(* CODESYS project getsystemtime.library
   DefaultNamespace: KOSTAL.AF2024.Core.GetSystemTime
   DocFormat: reStructuredText
   Description: Contains Functionalities to get the NT Real Time Clock
   Author: Frank Dümpelmann
   Title: KOSTAL.AF2024.Core.GetSystemTime
   Version: 1.0.1.0
   Company: KOSTAL GmbH & Co.KG
   Placeholder: KOSTAL.AF2024.Core.GetSystemTime

Project tree, tasks and I/O mapping:
  libraries: Tc2_Utilities, 3.3.47.0 (Beckhoff Automation GmbH); KOSTAL.AF2024.Core.System, 1.0.0.0 (KOSTAL GmbH & Co.KG)
  DUT/
    data type E_TIMESHIFT
    interface I_T_Timestruct: CopyTo, Day, DayOfWeek, Hour, iTimeStruct, Milliseconds, Minute, Month, Second, Year
    interface I_T_Timestruct_Owner: Day, DayOfWeek, Hour, Milliseconds, Minute, Month, Second, Timestruct, Year
    data type ST_TIMEZONE
    function block T_TIMESTRUCT [ST]: CopyTo, Day, DayOfWeek, Hour, iTimeStruct, Milliseconds, Minute, Month, Second, Timestruct, Year
  Interface/
    interface I_TimeSource: DateAndTime, GetTimeStruct, GetTimeZone, TimeStruct, Utc, Valid
  POU/
    function block FB_GetSystemTime [ST]: _formatTimeZone, amsNetId_timeServer, DateAndTime, FBmain, GetTimeStruct, GetTimeZone, Timeout, TimeStruct, Utc, Valid
  Project Information/
    function F_GetCompany [ST]
    function F_GetTitle [ST]
    function F_GetVersion [ST]
  Version/
    global variables Global_Version
*)

// DUT/E_TIMESHIFT
{attribute 'qualified_only'}
{attribute 'strict'}
TYPE E_TIMESHIFT :
(
	undef 		:= 0,
	positive 	:= 1,
	negative 	:= 2
);
END_TYPE

// DUT/ST_TIMEZONE
TYPE ST_TIMEZONE :
STRUCT
	timeshift	: E_TIMESHIFT;
	hours		: USINT;
	minutes		: USINT;
END_STRUCT
END_TYPE

// Version/Global_Version
{attribute 'TcGenerated'}
{attribute 'no-analysis'}
{attribute 'linkalways'}
// This function has been automatically generated from the project information.
VAR_GLOBAL CONSTANT
	{attribute 'const_non_replaced'}
	stLibVersion_KOSTAL_AF2024_Core_GetSystemTime : ST_LibVersion := (iMajor := 1, iMinor := 0, iBuild := 1, iRevision := 0, nFlags := 1, sVersion := '1.0.1.0');
END_VAR

// DUT/I_T_Timestruct
INTERFACE I_T_Timestruct EXTENDS KOSTAL_AF2024_Core_System.I_Interface

METHOD CopyTo
VAR_INPUT
	IN : REFERENCE TO Tc2_Utilities.TIMESTRUCT;
END_VAR
END_METHOD

PROPERTY PUBLIC Day : WORD
GET
END_GET
END_PROPERTY

PROPERTY PUBLIC DayOfWeek : WORD
GET
END_GET
END_PROPERTY

PROPERTY PUBLIC Hour : WORD
GET
END_GET
END_PROPERTY

PROPERTY iTimeStruct : Tc2_Utilities.TIMESTRUCT
GET
END_GET
END_PROPERTY

PROPERTY PUBLIC Milliseconds : WORD
GET
END_GET
END_PROPERTY

PROPERTY PUBLIC Minute : WORD
GET
END_GET
END_PROPERTY

PROPERTY PUBLIC Month : WORD
GET
END_GET
END_PROPERTY

PROPERTY PUBLIC Second : WORD
GET
END_GET
END_PROPERTY

PROPERTY PUBLIC Year : WORD
GET
END_GET
END_PROPERTY

END_INTERFACE

// DUT/I_T_Timestruct_Owner
INTERFACE I_T_Timestruct_Owner EXTENDS KOSTAL_AF2024_Core_System.I_Interface

PROPERTY PUBLIC Day : WORD
GET
END_GET
SET
END_SET
END_PROPERTY

PROPERTY PUBLIC DayOfWeek : WORD
GET
END_GET
SET
END_SET
END_PROPERTY

PROPERTY PUBLIC Hour : WORD
GET
END_GET
SET
END_SET
END_PROPERTY

PROPERTY PUBLIC Milliseconds : WORD
GET
END_GET
SET
END_SET
END_PROPERTY

PROPERTY PUBLIC Minute : WORD
GET
END_GET
SET
END_SET
END_PROPERTY

PROPERTY PUBLIC Month : WORD
GET
END_GET
SET
END_SET
END_PROPERTY

PROPERTY PUBLIC Second : WORD
GET
END_GET
SET
END_SET
END_PROPERTY

PROPERTY Timestruct : REFERENCE To Tc2_Utilities.TIMESTRUCT
GET
END_GET
END_PROPERTY

PROPERTY PUBLIC Year : WORD
GET
END_GET
SET
END_SET
END_PROPERTY

END_INTERFACE

// DUT/T_TIMESTRUCT
FUNCTION_BLOCK T_TIMESTRUCT IMPLEMENTS I_T_Timestruct, I_T_Timestruct_Owner
VAR
	_timestruct : Tc2_Utilities.TIMESTRUCT;
END_VAR

METHOD CopyTo
VAR_INPUT
	IN : REFERENCE TO Tc2_Utilities.TIMESTRUCT;
END_VAR

IN.wYear := _timestruct.wYear;
IN.wMonth := _timestruct.wMonth;
IN.wDay := _timestruct.wDay;
IN.wDayOfWeek := _timestruct.wDayOfWeek;
IN.wHour := _timestruct.wHour;
IN.wMinute := _timestruct.wMinute;
IN.wSecond := _timestruct.wSecond;
IN.wMilliseconds := _timestruct.wMilliseconds;
END_METHOD

PROPERTY PUBLIC Day : WORD
GET
Day := _timestruct.wDay;
END_GET
SET
_timestruct.wDay := Day;
END_SET
END_PROPERTY

PROPERTY PUBLIC DayOfWeek : WORD
GET
DayOfWeek := _timestruct.wDayOfWeek;
END_GET
SET
_timestruct.wDayOfWeek := DayOfWeek;
END_SET
END_PROPERTY

PROPERTY PUBLIC Hour : WORD
GET
Hour := _timestruct.wHour;
END_GET
SET
_timestruct.wHour := Hour;
END_SET
END_PROPERTY

PROPERTY iTimeStruct : Tc2_Utilities.TIMESTRUCT
GET
TimeStruct := _timestruct;
END_GET
END_PROPERTY

PROPERTY PUBLIC Milliseconds : WORD
GET
Milliseconds := _timestruct.wMilliseconds;
END_GET
SET
_timestruct.wMilliseconds := Milliseconds;
END_SET
END_PROPERTY

PROPERTY PUBLIC Minute : WORD
GET
Minute := _timestruct.wMinute;
END_GET
SET
_timestruct.wMinute := Minute;
END_SET
END_PROPERTY

PROPERTY PUBLIC Month : WORD
GET
Month := _timestruct.wMonth;
END_GET
SET
_timestruct.wMonth := Month;
END_SET
END_PROPERTY

PROPERTY PUBLIC Second : WORD
GET
Second := _timestruct.wSecond;
END_GET
SET
_timestruct.wSecond := Second;
END_SET
END_PROPERTY

PROPERTY Timestruct : REFERENCE To Tc2_Utilities.TIMESTRUCT
GET
Timestruct REF= _timestruct;
END_GET
END_PROPERTY

PROPERTY PUBLIC Year : WORD
GET
Year := _timestruct.wYear;
END_GET
SET
_timestruct.wYear := Year;
END_SET
END_PROPERTY

END_FUNCTION_BLOCK

// Interface/I_TimeSource
INTERFACE I_TimeSource EXTENDS KOSTAL_AF2024_Core_System.I_Interface

PROPERTY DateAndTime : DATE_AND_TIME
GET
END_GET
END_PROPERTY

METHOD PUBLIC GetTimeStruct : TIMESTRUCT
VAR_INPUT
END_VAR
END_METHOD

METHOD PUBLIC GetTimeZone : ST_TIMEZONE
VAR_INPUT
END_VAR
END_METHOD

(*
Description
===========
| Tc2_Utilities.TIMESTRUCT containing the current system time
*)
PROPERTY TimeStruct : I_T_Timestruct
GET
END_GET
END_PROPERTY

PROPERTY Utc : REFERENCE TO Tc2_Utilities.TIMESTRUCT
GET
END_GET
END_PROPERTY

(*
Description
===========
| Time source is valid
*)
PROPERTY Valid : BOOL
GET
END_GET
END_PROPERTY

END_INTERFACE

// POU/FB_GetSystemTime
(*

:Author: Frank Dümpelmann <f.duempelmann@kostal.com>, Martin Hundt <m.hundt@kostal.com>
:Date: 2018-11-19

Function
========
Reads windows system time and time zone


Usage notes
===============
| Asyncronous function block: FB_Main() method must be called cyclicly
| Implements interface I_Time

Methods and Properties
======================
| See bottom of this document for a detailed description of each method or property
| Methods starting with an underline(_) are internally used and can be ignored by the user

*)

FUNCTION_BLOCK FB_GetSystemTime IMPLEMENTS I_TimeSource

VAR
	_get_NT_Time	: Tc2_Utilities.NT_GetTime;	//Tc2_Utilities.NT_GetTime
	_getTimeZone	: Tc2_Utilities.FB_GetTimeZoneInformation;

	_amsNetId_timeServer	: STRING:= '';	//STRING:= '' - default local system
	_timeout	: TIME:= T#5S;	//TIME:= T#5s - default
	
	_TIMESTRUCT	: Tc2_Utilities.TIMESTRUCT;	//Tc2_Utilities.TIMESTRUCT
	_tTimestruct	: T_TIMESTRUCT;
	
	
	_dateAndTime	:	DATE_AND_TIME;
	_timezone		: ST_TIMEZONE;
	_timezoneBias	: DINT;
	
	_getUtc				: Tc2_Utilities.FB_TzSpecificLocalTimeToSystemTime;
	_UTC_TIMESTRUCT		: Tc2_Utilities.TIMESTRUCT;	//Tc2_Utilities.TIMESTRUCT
	
	_valid			: BOOL;	//BOOL
END_VAR

METHOD PROTECTED _formatTimeZone : ST_TIMEZONE;
VAR_INPUT
	timezoneBias	: DINT;
END_VAR

VAR
	_timezone	: ST_TIMEZONE;
	_biasAbs	: DINT;
	_minutes	: USINT;
	_hours		: USINT;
END_VAR
_biasAbs := ABS(timezoneBias);

IF timezoneBias > 0 THEN
	_timezone.timeshift := E_TIMESHIFT.negative;	//Negative Bias -> Positive Time zone
ELSE
	_timezone.timeshift := E_TIMESHIFT.positive;	
END_IF

_timezone.minutes  := DINT_TO_USINT(_biasAbs MOD 60);
_timezone.hours := DINT_TO_USINT((_biasAbs - _minutes)/60);


_formatTimeZone := _timezone;
END_METHOD

(*
Description
===========
| AMS NetID of  device to save log file to
| default: '' = Local device
*)
PROPERTY PUBLIC amsNetId_timeServer : STRING
GET

amsNetId_timeServer:= _amsNetId_timeServer;
END_GET
SET

_amsNetId_timeServer:= amsNetId_timeServer;
END_SET
END_PROPERTY

PROPERTY DateAndTime : DATE_AND_TIME
GET

DateAndTime:= _dateAndTime;
END_GET
END_PROPERTY

(*
Description
===========
| Main method, to be called cyclicly, e.g. in DeviceDefine
*)
METHOD PUBLIC FBmain
VAR_INPUT
END_VAR

IF NOT _get_NT_Time.START THEN 

	_get_NT_Time.START:= TRUE;
	
ELSIF _get_NT_Time.BUSY THEN 

	//wait

ELSIF _get_NT_Time.ERR THEN

	_get_NT_Time.START:= FALSE;
	_valid:= FALSE;
	
ELSIF NOT _getTimeZone.bExecute THEN 

	_getTimeZone.bExecute:= TRUE;
	
ELSIF _getTimeZone.bBusy THEN 

	//wait

ELSIF _getTimeZone.bError THEN

	 _getTimeZone.bExecute := FALSE;
	_valid:= FALSE;

ELSE
	//Valid -> Set output data
	_get_NT_Time.START:= FALSE;
	_getTimeZone.bExecute := FALSE;
	_valid:= TRUE;
	_TIMESTRUCT:= _get_NT_Time.TIMESTR;
	
	_tTimestruct.Timestruct := _TIMESTRUCT;
	
	_dateAndTime:= SYSTEMTIME_TO_DT(_get_NT_Time.TIMESTR);
	_timezoneBias := _getTimeZone.tzInfo.bias;
	_timezone 	:= _formatTimeZone(_timezoneBias);
	
END_IF

_get_NT_Time
	(
		NETID:= _amsNetId_timeServer, 
		START:= , 
		TMOUT:= _timeout, 

		BUSY		=> , 
		ERR			=> , 
		ERRID		=> , 
		TIMESTR	=> 
	);

	
_getTimeZone
	(
		sNETID:= _amsNetId_timeServer, 
		tTimeout:= _timeout, 
	);
	
_getUtc
	(	
		in:= _TIMESTRUCT, 
		tzInfo:= _getTimeZone.tzInfo, 
		out=> _UTC_TIMESTRUCT
	);
END_METHOD

METHOD PUBLIC GetTimeStruct : TIMESTRUCT
VAR_INPUT
END_VAR
getTimeStruct := _TIMESTRUCT;
END_METHOD

METHOD PUBLIC GetTimeZone : ST_TIMEZONE
VAR_INPUT
END_VAR
GetTimeZone := _timezone;
END_METHOD

(*
Description
===========
| Maximun execution time of block until fault is generated
*)
PROPERTY PUBLIC Timeout : TIME
GET

timeout:= _timeout;
END_GET
SET

_timeout:= timeout;
END_SET
END_PROPERTY

(*
Description
===========
| Tc2_Utilities.TIMESTRUCT containing the current system time
*)
PROPERTY TimeStruct : I_T_Timestruct
GET

TimeStruct := _tTimestruct;
END_GET
END_PROPERTY

PROPERTY Utc : REFERENCE TO Tc2_Utilities.TIMESTRUCT
GET

Utc	REF= _UTC_TIMESTRUCT;
END_GET
END_PROPERTY

(*
Description
===========
| Time source is valid
*)
PROPERTY Valid : BOOL
GET

Valid:= _valid;
END_GET
END_PROPERTY

END_FUNCTION_BLOCK

// Project Information/F_GetCompany
// This function has been automatically generated from the project information.
{attribute 'signature_flag' := '1073741824'}
{attribute 'TcGenerated'}
{attribute 'no-analysis'}
FUNCTION F_GetCompany : WSTRING
VAR_INPUT
	
END_VAR

F_GetCompany := "KOSTAL GmbH & Co.KG";

END_FUNCTION

// Project Information/F_GetTitle
// This function has been automatically generated from the project information.
{attribute 'signature_flag' := '1073741824'}
{attribute 'TcGenerated'}
{attribute 'no-analysis'}
FUNCTION F_GetTitle : WSTRING
VAR_INPUT
	
END_VAR

F_GetTitle := "KOSTAL.AF2024.Core.GetSystemTime";

END_FUNCTION

// Project Information/F_GetVersion
// This function has been automatically generated from the project information.
{attribute 'signature_flag' := '1073741824'}
{attribute 'TcGenerated'}
{attribute 'no-analysis'}
FUNCTION F_GetVersion : ST_LibVersion
VAR_INPUT
	
END_VAR

F_GetVersion.iMajor := 1;
F_GetVersion.iMinor := 0;
F_GetVersion.iBuild := 1;
F_GetVersion.iRevision := 0;
F_GetVersion.sVersion := '1.0.1.0';
F_GetVersion.nFlags := 1;

END_FUNCTION
